(* IEC 61131-3 sources: stdmachine/plc/src/02_Interfaces, 14 files *)

(* ---- I_AlarmSink.st ---- *)
// Réception des alarmes (docs/04 § 4, docs/14)
INTERFACE I_AlarmSink
METHOD Raise
VAR_INPUT
    nGlobalId : UDINT;
    nCode : UINT;
    nSubCode : UDINT;
    eSeverity : E_Severity;
END_VAR
END_METHOD
METHOD Clear
VAR_INPUT
    nGlobalId : UDINT;
    nCode : UINT;
END_VAR
END_METHOD
END_INTERFACE

(* ---- I_Beacon.st ---- *)
// Balise pilotée par le séquenceur auquel elle est rattachée (docs/02 § 8, docs/03 § 8.1)
INTERFACE I_Beacon
METHOD SetPattern
VAR_INPUT
    nPattern : UINT;             // bits de F_BeaconBits
    bBuzzer : BOOL;
END_VAR
END_METHOD
END_INTERFACE

(* ---- I_Group.st ---- *)
// Module : reçoit l'état agrégé de ses enfants, calculé par la station (docs/04 § 8)
INTERFACE I_Group
METHOD SetAggregate
VAR_INPUT
    eState : E_ObjState;
END_VAR
END_METHOD
END_INTERFACE

(* ---- I_InterlockProvider.st ---- *)
// Verrouillages d'une station (docs/04 § 4) : 0 si autorisé, sinon n° du verrouillage violé
INTERFACE I_InterlockProvider
METHOD Check : INT
VAR_INPUT
    nLocalId : UINT;
    nAction : UINT;
END_VAR
END_METHOD
END_INTERFACE

(* ---- I_Maintained.st ---- *)
// Compteurs de maintenance persistants d'un élément de pool (docs/11 § 5, D92) et leur restauration (docs/02 § 7.4)
INTERFACE I_Maintained
// Objet du projet auquel appartiennent les compteurs (persistant : survit au redémarrage du PLC)
PROPERTY StableId : UDINT
GET
END_GET
END_PROPERTY
PROPERTY ActionCount : UDINT
GET
END_GET
END_PROPERTY
PROPERTY ErrorCount : UDINT
GET
END_GET
END_PROPERTY
PROPERTY MotionHours : LREAL
GET
END_GET
END_PROPERTY
METHOD RestoreCounters
VAR_INPUT
    nActions : UDINT;
    nErrors : UDINT;
    fHours : LREAL;
END_VAR
END_METHOD
END_INTERFACE

(* ---- I_ManualHost.st ---- *)
// Ce que le canal manuel lit de son hôte : une station, ou la machine pour le canal 0 (docs/05 § 7)
INTERFACE I_ManualHost
// Objet de n° local nLocalId, 0 si absent
METHOD ObjectAt : I_Object
VAR_INPUT
    nLocalId : UINT;
END_VAR
END_METHOD
// Position nommée à apprendre, 0 si l'hôte n'en a pas (la machine n'a pas de positions nommées)
METHOD NamedPos : POINTER TO ST_NamedPos
VAR_INPUT
    nIndex : INT;
END_VAR
END_METHOD
PROPERTY State : E_State
GET
END_GET
END_PROPERTY
PROPERTY Mode : E_Mode
GET
END_GET
END_PROPERTY
END_INTERFACE

(* ---- I_MoverMotion.st ---- *)
// Mouvement d'un mover hors process (mode manuel, docs/05 § 6.5) : le gestionnaire de movers tient l'occupation
// à jour. Donnée aux objets Mover par GVL_IoRef.ipMovers.
INTERFACE I_MoverMotion
// Déplacement vers une position quelconque du plan ; fSpeedPct en % de la vitesse par défaut des movers
METHOD MoveFree : BOOL
VAR_INPUT
    nMover : USINT;
    stPos : ST_Position;
    fSpeedPct : LREAL;
END_VAR
END_METHOD
METHOD StopMover
VAR_INPUT
    nMover : USINT;
END_VAR
END_METHOD
METHOD Moving : BOOL
VAR_INPUT
    nMover : USINT;
END_VAR
END_METHOD
METHOD Position : ST_Position
VAR_INPUT
    nMover : USINT;
END_VAR
END_METHOD
END_INTERFACE

(* ---- I_Node.st ---- *)
// Tout ce qui porte un override et un état : machine, station, module, objet (docs/04 § 4)
INTERFACE I_Node
PROPERTY EffectiveOverride : LREAL
GET
END_GET
END_PROPERTY
PROPERTY NodeState : E_ObjState
GET
END_GET
END_PROPERTY
END_INTERFACE

(* ---- I_Object.st ---- *)
// Contrat de tout objet (docs/04 § 4)
INTERFACE I_Object EXTENDS I_Node
METHOD Configure : BOOL
VAR_INPUT
    refCfg : REFERENCE TO ST_ObjConfig;
    nStation : UINT;             // 0 = machine (D92 : le n° de station n'est pas dans ST_ObjConfig)
    nPoolIndex : UINT;
    ipParent : I_Node;
    ipLocks : I_InterlockProvider;
    ipAlarms : I_AlarmSink;
END_VAR
END_METHOD
METHOD Start : E_StartResult
VAR_INPUT
    nAction : UINT;
    refParams : REFERENCE TO ST_ActParams;
    bManual : BOOL;
END_VAR
END_METHOD
METHOD Abort
END_METHOD
METHOD Ack : BOOL
END_METHOD
METHOD Cycle
END_METHOD
METHOD ForceInput
VAR_INPUT
    nSignal : USINT;             // S1..S8 ; 0 = rendre la main à la simulation
    fValue : LREAL;
END_VAR
END_METHOD
PROPERTY Info : REFERENCE TO ST_ObjectInfo
GET
END_GET
END_PROPERTY
PROPERTY ActStatus : E_ActStatus
GET
END_GET
END_PROPERTY
PROPERTY Results : REFERENCE TO ST_ActResults
GET
END_GET
END_PROPERTY
PROPERTY Status : REFERENCE TO ST_ObjStatus
GET
END_GET
END_PROPERTY
END_INTERFACE

(* ---- I_ObjectHost.st ---- *)
// Registre d'objets d'une station ou de la machine (docs/04 § 9), rempli par FB_ObjectFactory
INTERFACE I_ObjectHost
METHOD ClearObjects
END_METHOD
METHOD SetObject
VAR_INPUT
    nLocalId : UINT;
    ipObj : I_Object;
END_VAR
END_METHOD
END_INTERFACE

(* ---- I_ObjectPools.st ---- *)
// Pools d'objets (docs/04 § 9) : instances déclarées une fois pour toutes, attribuées au déploiement par
// FB_ObjectFactory. La bibliothèque fournit FB_DefaultPools ; un projet peut donner les siens.
INTERFACE I_ObjectPools
// Nombre d'éléments du pool d'un type, 0 = type absent
METHOD PoolSize : UINT
VAR_INPUT
    nType : UINT;
END_VAR
END_METHOD
// N° du pool d'un type : deux types qui partagent un pool (axe linéaire et rotatif, modules) ont le même n°
METHOD PoolId : UINT
VAR_INPUT
    nType : UINT;
END_VAR
END_METHOD
// Élément nIndex (1..PoolSize) du pool d'un type
METHOD Element : I_Object
VAR_INPUT
    nType : UINT;
    nIndex : UINT;
END_VAR
END_METHOD
END_INTERFACE

(* ---- I_OrderAware.st ---- *)
// Objet qui réagit au changement d'OF (compteur, P3 : remise à zéro au changement d'OF, docs/03 § 8.4)
INTERFACE I_OrderAware
METHOD OnOrderChange
END_METHOD
END_INTERFACE

(* ---- I_PlanarDriver.st ---- *)
// Pilote du système planaire (docs/05 § 6). Le séquenceur ne donne que des destinations ; trajets et évitement
// de collision sont faits par le système planaire. FB_PlanarSim l'implémente en simulation ; le pilote Tc3 Planar
// (projet de la machine ou bibliothèque à venir) implémente la même interface.
INTERFACE I_PlanarDriver
METHOD Activate : BOOL              // TRUE quand le système est actif
VAR_INPUT
    bEnable : BOOL;
END_VAR
END_METHOD
METHOD MoveTo : BOOL                // TRUE si la commande est acceptée
VAR_INPUT
    nMover : USINT;
    stPos : ST_Position;
    fVelocity : LREAL;               // mm/s, override déjà appliqué par le pilote
    fAcceleration : LREAL;
END_VAR
END_METHOD
METHOD StopAll
END_METHOD
METHOD StopMover                    // arrêt contrôlé d'un mover (mode manuel)
VAR_INPUT
    nMover : USINT;
END_VAR
END_METHOD
METHOD AckError
END_METHOD
METHOD Cycle
VAR_INPUT
    fOverride : LREAL;               // override machine effectif, %
END_VAR
END_METHOD
METHOD MoverPosition : ST_Position
VAR_INPUT
    nMover : USINT;
END_VAR
END_METHOD
METHOD MoverMoving : BOOL
VAR_INPUT
    nMover : USINT;
END_VAR
END_METHOD
METHOD MoverDetected : BOOL
VAR_INPUT
    nMover : USINT;
END_VAR
END_METHOD
METHOD SetInitialPosition           // simulation : poser un mover sur le plan
VAR_INPUT
    nMover : USINT;
    stPos : ST_Position;
END_VAR
END_METHOD
PROPERTY Active : BOOL
GET
END_GET
END_PROPERTY
PROPERTY ErrorCode : UINT          // 0 ou erreur du type Système planaire (100 collision, 101 mover non détecté, 102 groupe)
GET
END_GET
END_PROPERTY
PROPERTY ErrorSubCode : UDINT
GET
END_GET
END_PROPERTY
END_INTERFACE

(* ---- I_SafetyCircuits.st ---- *)
// Objet Sécurités : la station (ou la machine) lit l'état de ses circuits (docs/03 § 8.2, docs/05 § 4.2)
INTERFACE I_SafetyCircuits
PROPERTY AllOk : BOOL
GET
END_GET
END_PROPERTY
END_INTERFACE
